TYPE "ST_AirPressureOutImm"
VERSION : 0.1
   STRUCT
      "LowPressure" : Bool;
      "OperatingPressure" : Bool;
      "PressureOk" : Bool;
      "Contradictory" : Bool;
      "Quality" : Bool;
   END_STRUCT;
END_TYPE
